(* IEC 61131-3 sources: nautilus/sparkplug/host/codegen/testdata, 1 file *)

(* ---- sparkplug_types.st ---- *)
(*
  Generated by `nautilus sparkplug import` from the group's NBIRTH template
  definitions. Do not edit — re-run the import when a site's UDTs change.
  Group: PomonaWRD
*)

TYPE
  Motor : STRUCT
    Speed : LREAL;
    Run : BOOL;
  END_STRUCT;
  Skid : STRUCT
    Main : Motor;
    Hours : DINT;
  END_STRUCT;
END_TYPE

(* Add the tags your program uses to its VAR_EXTERNAL block. The __Online,
   __LastBirthMs and __Rebirth tags are synthesized by the driver: interlock
   on __Online before trusting a site's values, and pulse __Rebirth to force
   a resync.

VAR_EXTERNAL
  W6_PLC1_Pump_Run : BOOL;
  W6_PLC1_Pump_SpeedSP : LREAL;
  W6_PLC1__Online : BOOL;
  W6_Pump1 : Motor;
  W6_Pump1_Speed : LREAL;
  W6_Site_Name : STRING;
  W6_Skid_A : Skid;
  W6_Skid_A_Main_Run : BOOL;
  W6_Well_LastSample : LINT;
  W6_Well_Level : LREAL;
  W6__LastBirthMs : LINT;
  W6__Online : BOOL;
  W6__Rebirth : BOOL;
  W7_Pump1 : Motor;
  W7_Pump1_Speed : LREAL;
  W7_Well_Level : LREAL;
  W7__LastBirthMs : LINT;
  W7__Online : BOOL;
  W7__Rebirth : BOOL;
END_VAR
*)
